// TIA Portal V21 export
// export: Created 2026-11-11T00:48:18.830974Z, ExportSetting WithDefaults, DisplayName Totally Integrated Automation Portal, DisplayVersion V21 Update 3, DisplayName STEP 7 Professional, DisplayVersion V21 Update 3, DisplayName STEP 7 Safety, DisplayVersion V21, DisplayName Tech WebApplication, DisplayVersion V21, DisplayName WinCC Basic/Comfort/Advanced, DisplayVersion V21 Update 3, DisplayName WinCC Unified, DisplayVersion V21 Update 3
FUNCTION_BLOCK "FB_Scl_sl059"   // FB34, SCL
{ S7_Optimized_Access := 'TRUE' }
VERSION : 0.1
// stored: AutoNumber true, IsIECCheckEnabled false, IsRetainMemResEnabled false, MemoryReserve 100, SetENOAutomatically false, UDAEnableTagReadback false
   VAR_INPUT
      v_area_src : Byte;
      v_dbnumber_src : DInt;
      v_byteoffset_src : DInt;
      v_area_dest : Byte;
      v_dbnumber_dest : DInt;
      v_byteoffset_dest : DInt;
      v_count : DInt;
   END_VAR
BEGIN
   POKE_BLK(area_src := #v_area_src, dbNumber_src := #v_dbnumber_src, byteOffset_src := #v_byteoffset_src, area_dest := #v_area_dest, dbNumber_dest := #v_dbnumber_dest, byteOffset_dest := #v_byteoffset_dest, count := #v_count);
END_FUNCTION_BLOCK
